DATA_BLOCK "GDB_ProfileCases"
{ S7_Optimized_Access := 'TRUE' }
VERSION : 0.1
NON_RETAIN
VAR
    Complete {ExternalWritable := 'False'} : Bool;
    Count {ExternalWritable := 'False'} : Int;
    Passed {ExternalWritable := 'False'} : Array[1..57] of Bool;
END_VAR
BEGIN
END_DATA_BLOCK
